(* PLC project Vn_and3_edit_pin_removed, Beckhoff Automation GmbH TwinCAT PLC Control 3.5.13.21 *)
(* stored: creationDateTime 1970-01-01T00:00:00 *)

PROGRAM Vn_and3_edit_pin_removed

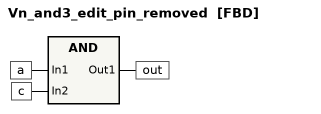
(* FBD diagram, written out as Structured Text *)
out := a AND c;
END_PROGRAM
